TYPE "ST_PressDemoOutCmd"
VERSION : 0.1
   STRUCT
      "CycleCompleted" : Bool;
   END_STRUCT;
END_TYPE
